Fanuc KAREL source: kt00124.KL

-- PROVISIONAL review KL for V1013-1; original PC SHA256 542998c237c209d3e7366fa9db1205813e718735746e1ec3ff2c3be07451af29
-- Incomplete behavior may be omitted. Consult companion uncertainty JSON. Do not deploy.
PROGRAM KT00124
%NOLOCKGROUP
VAR
  R2 : REAL
  OUT : REAL
-- UNRESOLVED_DECL H1 type=002017
BEGIN
  -- UNRESOLVED_PC offsets 5-19; opcodes 2E,22,9D,33,B4
  -- UNRESOLVED_PC offsets 24-35; opcodes 2E,23
  -- UNRESOLVED_PC offsets 40-65; opcodes 22,9D,33,B3,21,29,64,29,6C,23
  -- UNRESOLVED_PC offsets 70-74; opcodes 7F
END KT00124
